// TwinCAT 3 PLC project DriveStateTests
// ProgramVersion: 3.1.4026.22
// libraries:
//   Tc2_Standard, * (Beckhoff Automation GmbH)
//   Tc2_System, * (Beckhoff Automation GmbH)
// project tree:
//   StateMachineControl/DUTs/ E_DriveState.TcDUT
//   StateMachineControl/POUs/ F_DecodeDriveState.TcPOU, FB_StateMachineControl.TcPOU
//   StateMachineControl/tests/POUs/ PRG_DriveStateTests.TcPOU
//   StateMachineControl/tests/ DriveStateTestTask.TcTTO
// (motion and I/O tree: see PLC project experimentsequencertests)
// real-time tasks:
//   TASK DriveStateTestTask: cycle T#10ms, priority 1, ADS port 350
//   TASK TestTask: cycle T#10ms, priority 2, ADS port 351

CONFIGURATION DriveStateTests
    RESOURCE PLC ON TwinCAT3
        TASK DriveStateTestTask(INTERVAL := T#10ms, PRIORITY := 1);
        PROGRAM PRG_DriveStateTests WITH DriveStateTestTask : PRG_DriveStateTests;
    END_RESOURCE
END_CONFIGURATION

// ---- StateMachineControl/DUTs/E_DriveState.TcDUT
{attribute 'qualified_only'}
{attribute 'strict'}
{attribute 'to_string'}
TYPE E_DriveState :
(
    UNKNOWN := 0,

    // CiA402 "Switch on disabled"
    SWITCH_ON_DISABLED := 10,

    // CiA402 "Ready to switch on"
    READY_TO_SWITCH_ON := 20,

    // CiA402 "Switched on"
    SWITCHED_ON := 30,

    // CiA402 "Operation enabled"
    OPERATION_ENABLED := 40,

    // CiA402 "Fault"
    FAULT := 90
);
END_TYPE

// ---- StateMachineControl/tests/POUs/PRG_DriveStateTests.TcPOU
PROGRAM PRG_DriveStateTests
VAR
    driveControl : FB_StateMachineControl;
    testsExecuted : BOOL := FALSE;
    testsPassed : BOOL := FALSE;
    failureCount : UDINT := 0;
END_VAR

IF NOT testsExecuted THEN
    (* Decoder must ignore manufacturer/status bits outside the CiA402 mask. *)
    IF F_DecodeDriveState(16#0060) <> E_DriveState.SWITCH_ON_DISABLED
        OR F_DecodeDriveState(16#00E0) <> E_DriveState.SWITCH_ON_DISABLED
        OR F_DecodeDriveState(16#0021) <> E_DriveState.READY_TO_SWITCH_ON
        OR F_DecodeDriveState(16#0023) <> E_DriveState.SWITCHED_ON
        OR F_DecodeDriveState(16#0027) <> E_DriveState.OPERATION_ENABLED
        OR F_DecodeDriveState(16#0008) <> E_DriveState.FAULT
        OR F_DecodeDriveState(16#0000) <> E_DriveState.UNKNOWN THEN
        failureCount := failureCount + 1;
    END_IF

    driveControl(statusWord := 16#0027, enable := FALSE);
    IF driveControl.controlWord <> 16#0000 THEN failureCount := failureCount + 1; END_IF

    driveControl(statusWord := 16#0060, enable := TRUE);
    IF driveControl.controlWord <> 16#0006 THEN failureCount := failureCount + 1; END_IF
    driveControl(statusWord := 16#0021, enable := TRUE);
    IF driveControl.controlWord <> 16#0007 THEN failureCount := failureCount + 1; END_IF
    driveControl(statusWord := 16#0023, enable := TRUE);
    IF driveControl.controlWord <> 16#000F THEN failureCount := failureCount + 1; END_IF
    driveControl(statusWord := 16#0027, enable := TRUE);
    IF driveControl.controlWord <> 16#000F THEN failureCount := failureCount + 1; END_IF

    (* Fault reset is exactly one call while the fault remains asserted. *)
    driveControl(statusWord := 16#0008, enable := TRUE);
    IF driveControl.controlWord <> 16#0080 THEN failureCount := failureCount + 1; END_IF
    driveControl(statusWord := 16#0008, enable := TRUE);
    IF driveControl.controlWord <> 16#0000 THEN failureCount := failureCount + 1; END_IF
    driveControl(statusWord := 16#0060, enable := TRUE);
    driveControl(statusWord := 16#0008, enable := TRUE);
    IF driveControl.controlWord <> 16#0080 THEN failureCount := failureCount + 1; END_IF

    (* UNKNOWN converges with the safe shutdown command. *)
    driveControl(statusWord := 16#0000, enable := TRUE);
    IF driveControl.driveState <> E_DriveState.UNKNOWN OR driveControl.controlWord <> 16#0006 THEN
        failureCount := failureCount + 1;
    END_IF

    testsExecuted := TRUE;
    testsPassed := (failureCount = 0);
END_IF

END_PROGRAM

// ---- StateMachineControl/POUs/FB_StateMachineControl.TcPOU
FUNCTION_BLOCK FB_StateMachineControl
VAR_INPUT
    statusWord : UINT; // 0x6041
    enable      : BOOL := TRUE;
END_VAR
VAR_OUTPUT
    controlWord : UINT;      // 0x6040
    driveState   : E_DriveState;
END_VAR
VAR
    faultResetPulsed : BOOL := FALSE;
END_VAR
VAR CONSTANT
    // Common CiA402 control commands (0x6040)
    CW_DISABLE_VOLTAGE : UINT := 16#0000;
    CW_SHUTDOWN        : UINT := 16#0006;
    CW_SWITCH_ON       : UINT := 16#0007;
    CW_ENABLE_OP       : UINT := 16#000F;
    CW_FAULT_RESET     : UINT := 16#0080;
END_VAR

driveState := F_DecodeDriveState(statusWord);

// Disable requested: force safe output
IF NOT enable THEN
    controlWord := CW_DISABLE_VOLTAGE;
    faultResetPulsed := FALSE;
    RETURN;
END_IF

CASE driveState OF

    E_DriveState.FAULT:
        // Fault reset should be a pulse. One scan is usually enough.
        IF NOT faultResetPulsed THEN
            controlWord := CW_FAULT_RESET;
            faultResetPulsed := TRUE;
        ELSE
            controlWord := CW_DISABLE_VOLTAGE;
        END_IF

    E_DriveState.SWITCH_ON_DISABLED:
        controlWord := CW_SHUTDOWN;
        faultResetPulsed := FALSE;

    E_DriveState.READY_TO_SWITCH_ON:
        controlWord := CW_SWITCH_ON;
        faultResetPulsed := FALSE;

    E_DriveState.SWITCHED_ON:
        controlWord := CW_ENABLE_OP;
        faultResetPulsed := FALSE;

    E_DriveState.OPERATION_ENABLED:
        controlWord := CW_ENABLE_OP;
        faultResetPulsed := FALSE;

    ELSE
        // UNKNOWN: converge from below (safe)
        controlWord := CW_SHUTDOWN;
        faultResetPulsed := FALSE;
END_CASE

END_FUNCTION_BLOCK

// ---- StateMachineControl/POUs/F_DecodeDriveState.TcPOU
FUNCTION F_DecodeDriveState : E_DriveState
VAR_INPUT
    statusWord : UINT; // 0x6041
END_VAR
VAR
    masked : UINT;
END_VAR

masked := statusWord AND 16#006F;

IF (masked AND 16#0008) <> 0 THEN
    // bit3 = Fault
    F_DecodeDriveState := E_DriveState.FAULT;
ELSIF masked = 16#0060 THEN
    // Switch on disabled
    F_DecodeDriveState := E_DriveState.SWITCH_ON_DISABLED;
ELSIF masked = 16#0021 THEN
    // Ready to switch on
    F_DecodeDriveState := E_DriveState.READY_TO_SWITCH_ON;
ELSIF masked = 16#0023 THEN
    // Switched on
    F_DecodeDriveState := E_DriveState.SWITCHED_ON;
ELSIF masked = 16#0027 THEN
    // Operation enabled
    F_DecodeDriveState := E_DriveState.OPERATION_ENABLED;
ELSE
    F_DecodeDriveState := E_DriveState.UNKNOWN;
END_IF

END_FUNCTION
